{region 'Documentation'}
(*!
<summary>Checks that the rising-edge count is greater than or equal to the minimum.</summary>
<description>

Observation and accumulated-count handling come from AssertionEdgeCountBase. Evaluate
checks the held count independently of Enable; reset clears the count and baseline.

</description>
*)
{endregion}
FUNCTION_BLOCK AssertRisingEdgeCntGreaterEqual EXTENDS AssertionEdgeCountBase
VAR_INPUT
    Minimum : UINT; //! Inclusive lower bound of the comparison; for a range, must not exceed Maximum.
END_VAR

SUPER^();

{region 'Documentation'}
(*!
<summary>Observe through the base, then evaluate the count with Error priority.</summary>
*)
{endregion}
METHOD PROTECTED Assert
VAR
    Message : STRING(GVL_Constants.MessageLength);
    MinimumText : STRING(GVL_Constants.AssertionValueLength);
    ActualText : STRING(GVL_Constants.AssertionValueLength);
END_VAR
SUPER^.Assert();

IF NOT EvaluationActive THEN
    RETURN;
END_IF;

IF Result = E_Result.Error THEN
    RETURN;
END_IF;

IF Result = E_Result.Failed THEN
    RETURN;
END_IF;

IF EdgeCount < Minimum THEN
    MinimumText := UINT_TO_STRING(Minimum);
    ActualText := UINT_TO_STRING(EdgeCount);
    Message := CONCAT('Assertion failed: rising edge count is below minimum. Minimum = ',
        MinimumText);
    Message := CONCAT(Message, ', Actual = ');
    Message := CONCAT(Message, ActualText);
    Message := CONCAT(Message, '.');
    Fail(Message := Message);
    RETURN;
END_IF;

Pass();
END_METHOD

{region 'Documentation'}
(*!
<summary>Recognize a rising edge without changing observation state.</summary>
*)
{endregion}
METHOD PROTECTED IsMatchingEdge : BOOL //! TRUE when PreviousValue and CurrentValue form the edge selected by this Assertion.
VAR_INPUT
    PreviousValue : BOOL; //! Signal value from the preceding active observation.
    CurrentValue : BOOL; //! Signal value from the current active observation.
END_VAR
IsMatchingEdge := NOT PreviousValue AND CurrentValue;
END_METHOD

END_FUNCTION_BLOCK

(* stored: Version 1.1.0.1
   POU AssertRisingEdgeCntGreaterEqual: Id {dac7fb03-3d01-4fa3-9d2f-15bbf7435bec}, SpecialFunc None
   Folder Internal: Id {7ec32089-4f9b-4230-b98a-9ee5624c1526}
   Method Assert: Id {647491af-2ce4-40e1-b9d9-8b29a1a43116}
   Method IsMatchingEdge: Id {a00d823d-ff79-4101-a246-683d63f15128} *)
